(* IEC 61131-3 sources: kns-port-domestic/tools/port_metrics_tests/fixtures/app/src/DUTs, 2 files *)

(* ---- E_PumpMode.dut.st ---- *)
{attribute 'qualified_only'}
{attribute 'strict'}
TYPE E_PumpMode :
(
    Auto := 1,
    Manual := 2
) UINT;
END_TYPE

(* ---- ST_PumpCfg.dut.st ---- *)
TYPE ST_PumpCfg :
STRUCT
    rSpeedMax_Hz : REAL := 50.0; // предел частоты
    tStartDelay : TIME := T#5S;
END_STRUCT
END_TYPE
